{attribute 'qualified_only'}
VAR_GLOBAL
	
	// BistableSingleCoilRelay ToggleVirtualState
	// Manually toggle internal, virtual relay state when mismatch with real, physical	
	Shutter1OpenRelayToggle : BOOL := FALSE;
	Shutter1CloseRelayToggle : BOOL := FALSE;
	
	// Shutters
	Shutter1Cmd : stShutterCommand;
	Shutter1CmdExecute : BOOL := FALSE;
	Shutter1Position : stShutterPosition;
    Shutter1State : eShutterStateType;
	ShutterUpSavedPos : stShutterPosition;
	ShutterDownSavedPos : stShutterPosition;

END_VAR

(* stored: Version 1.1.0.1
   GVL gvlHA: Id {0181db7e-994c-475a-978f-c286ac6dc635} *)
